(* IEC 61131-3 sources: Lasal-MCP/examples/SampleSource/LASALScreenAdvancedSolution/LASALScreenAdvancedSolution/LASALScreenAdvacnedSolution/Stations/Terminal/HMI/Class/DataRecordFileRead, 1 file *)

(* ---- DataRecordFileRead.st ---- *)
(*!
<Class
	Name               = "DataRecordFileRead"
	Revision           = "0.0"
	RealtimeTask       = "false"
	CyclicTask         = "false"
	BackgroundTask     = "true"
	DefBackground      = "10 ms"
	Sigmatek           = "false"
	OSInterface        = "false"
	HighPriority       = "false"
	Automatic          = "false"
	UpdateMode         = "Prescan"
	SharedCommandTable = "true"
	Objectsize         = "(444,120)">
	<Channels>
		<Server Name="IntError" Visualized="false" Initialize="false" WriteProtected="true" Retentive="false"/>
		<Server Name="ReadStep" Visualized="false" Initialize="false" WriteProtected="true" Retentive="false"/>
		<Server Name="StartRead" Visualized="true" Initialize="false" WriteProtected="false" Retentive="false"/>
		<Client Name="_FileSys" Required="false" Internal="false"/>
		<Client Name="_StdLib" Required="false" Internal="false"/>
		<Client Name="StringRAM" Required="true" Internal="false"/>
	</Channels>
</Class>
*)
DataRecordFileRead : CLASS
	TYPE
	  _READ_STEPS :  //! <Type Public="true" Name="_READ_STEPS"/>
	  (
	    RS_Idle,
	    RS_GetFileName,
	    RS_Open,
	    RS_WaitFileOpen,
	    RS_GetLength,
	    RS_WaitForGetLength,
	    RS_ReadFile,
	    RS_WaitForReadFile,
	    RS_CloseFile,
	    RS_WaitForClose,
	    RS_Error
	  )$UDINT;
	END_TYPE
  //Servers:
	ReadStep 	: SvrChCmd__READ_STEPS_PTofCls_DataRecordFileRead;
	IntError 	: SvrCh_DINT;
	StartRead 	: SvrCh_DINT;
  //Clients:
	_FileSys 	: CltChCmd__FileSys;
	_StdLib 	: CltChCmd__StdLib;
	StringRAM 	: CltChCmd_StringRAM;
  //Variables:
		FileName : ARRAY [0..99] OF CHAR;

		AsyncId 	: DINT;
		FileHandle 	: DINT;
		FileLength 	: UDINT;
		pReadData 	: ^DINT;
		FileIsRead 	: BOOL;
  //Functions:

	FUNCTION VIRTUAL GLOBAL Background
		VAR_INPUT
			EAX 	: UDINT;
		END_VAR
		VAR_OUTPUT
			state (EAX) 	: UDINT;
		END_VAR;

	FUNCTION GLOBAL ReadKoords
		VAR_INPUT
			pNoOfCoordinates 	: ^UDINT;
		END_VAR
		VAR_OUTPUT
			pCoord 	: ^_DOT;
		END_VAR;

	FUNCTION GLOBAL GetReadState
		VAR_OUTPUT
			IsRead 	: BOOL;
		END_VAR;

	FUNCTION GLOBAL SetReadState
		VAR_INPUT
			IsDrawing 	: BOOL;
		END_VAR;

	FUNCTION GLOBAL StartReading
		VAR_INPUT
			BufferSize 	: UDINT;
		END_VAR;
  //Tables:
	FUNCTION @STD
		VAR_OUTPUT
			ret_code	: CONFSTATES;
		END_VAR;
	FUNCTION GLOBAL TAB @CT_;
END_CLASS;

#pragma usingLtd _FileSys
#pragma usingLtd _StdLib
#pragma usingLtd StringRAM

FUNCTION VIRTUAL GLOBAL DataRecordFileRead::Background
	VAR_INPUT
		EAX 	: UDINT;
	END_VAR
	VAR_OUTPUT
		state (EAX) 	: UDINT;
	END_VAR
  VAR
  	stringLength : UDINT;
    asyncState : DINT;
    length : UDINT;
  END_VAR

  // ==========================================================================
  case ReadStep of

    // --------------------------------------------------------------
  	RS_Idle:

      if (StartRead = 1) then
         StartRead := 0;

         ReadStep := RS_GetFileName;
      end_if;

    // --------------------------------------------------------------
  	RS_GetFileName:

      stringLength := StringRAM.GetLength();

      StringRAM.GetDataAt(pData:= #FileName[0],
                          udSize:= stringLength,
                          udAt:= 0);

      ReadStep := RS_Open;

    // --------------------------------------------------------------
  	RS_Open:

      AsyncId := _FileSys.FileOpen_A(Async:= 1,
                                     filename:= #FileName[0],
                                     attributes:= ATT_READ_WRITE);

      ReadStep := RS_WaitFileOpen;

    // --------------------------------------------------------------
  	RS_WaitFileOpen:

      asyncState := _FileSys.GetAsyncState(ID:= to_udint(AsyncId),
                                           Erg:= #FileHandle);

      // ==================================================
      case asyncState of
        //---------------------------------------
        0:
          if (FileHandle >= 0) then
              ReadStep := RS_GetLength;
          else
            IntError := -1;
            ReadStep := RS_Error;
          end_if;

        //---------------------------------------
        RT_ERG_DELETED,
        RT_INVALID_ID:
          IntError := -2;
          ReadStep := RS_Error;

        //---------------------------------------
        RT_NOT_STARTED,
        RT_IN_PROGRESS:

      end_case;
      // ==================================================

    // --------------------------------------------------------------
  	RS_GetLength:

      AsyncId := _FileSys.FileLength_A(Async:= 1,
                                       handle:= FileHandle);
      ReadStep := RS_WaitForGetLength;

    // --------------------------------------------------------------
  	RS_WaitForGetLength:

      asyncState := _FileSys.GetAsyncState(ID:= to_udint(AsyncId),
                                           Erg:= #FileLength$dint);
        // ==================================================
      case asyncState of
        //---------------------------------------
        0:
          if (FileLength >= 0) then
            ReadStep := RS_ReadFile;
          end_if;

        //---------------------------------------
        RT_ERG_DELETED,
        RT_INVALID_ID:
            IntError := -3;
            ReadStep := RS_Error;

        //---------------------------------------
        RT_NOT_STARTED,
        RT_IN_PROGRESS:

      end_case;
     // ==================================================

    // --------------------------------------------------------------
  	RS_ReadFile:

      if (pReadData <> NIL) then
        _StdLib.Free(mptr:=pReadData);
      end_if;

      pReadData$^void := oc_StdLib.Malloc(size:= FileLength);

      AsyncId$UDINT := _FileSys.FileRead_A(Async:= 1,
                                           handle:= FileHandle,
                                           buffer:= pReadData,
                                           length:= FileLength);
      ReadStep := RS_WaitForReadFile;

    // --------------------------------------------------------------
  	RS_WaitForReadFile:

      asyncState := _FileSys.GetAsyncState(ID:= to_udint(AsyncId),
                                           Erg:= #FileHandle);
      // ==================================================
      case asyncState of
        //---------------------------------------
        0:
          if (length <> FileLength) then
            ReadStep := RS_CloseFile;
          else
            IntError := -4;
            ReadStep := RS_Error;
          end_if;

        //---------------------------------------
        RT_ERG_DELETED,
        RT_INVALID_ID:
          IntError := -5;
          ReadStep := RS_Error;

        //---------------------------------------
        RT_NOT_STARTED,
        RT_IN_PROGRESS:

        end_case;
       // ==================================================

    // --------------------------------------------------------------
  	RS_CloseFile:

      AsyncId := _FileSys.FileClose_A(Async:= 1,
                                      handle:= FileHandle);

      ReadStep := RS_WaitForClose;

    // --------------------------------------------------------------
  	RS_WaitForClose:

     asyncState := _FileSys.GetAsyncState(ID:= to_udint(AsyncId),
                                          Erg:= #FileHandle);

      // ==================================================
      case asyncState of
        //---------------------------------------
        0:
          if (FileHandle >= 0) then
            FileIsRead := TRUE;
            ReadStep := RS_Idle;
          else
            IntError := -6;
            ReadStep := RS_Error;
          end_if;
      end_case;
      // ==================================================

    // --------------------------------------------------------------
  	RS_Error:

  end_case;
  // ==========================================================================

	state := READY;

END_FUNCTION

FUNCTION GLOBAL DataRecordFileRead::ReadKoords
	VAR_INPUT
		pNoOfCoordinates 	: ^UDINT;
	END_VAR
	VAR_OUTPUT
		pCoord 	: ^_DOT;
	END_VAR

  pNoOfCoordinates^ := FileLength;
  pCoord := pReadData$^_DOT;

END_FUNCTION

FUNCTION GLOBAL DataRecordFileRead::GetReadState
	VAR_OUTPUT
		IsRead 	: BOOL;
	END_VAR

  IsRead := FileIsRead;

END_FUNCTION

FUNCTION GLOBAL DataRecordFileRead::SetReadState
	VAR_INPUT
		IsDrawing 	: BOOL;
	END_VAR

  FileIsRead := IsDrawing;

END_FUNCTION

FUNCTION GLOBAL DataRecordFileRead::StartReading
	VAR_INPUT
		BufferSize 	: UDINT;
	END_VAR

  if (pReadData <> NIL) then
    _StdLib.Free(mptr:=pReadData);
  end_if;

  pReadData$^void := _StdLib.Malloc(size:=BufferSize);

  if (pReadData <> NIL) then
      _StdLib.MemSet(dest:= pReadData,
                     value:= 0,
                     size:= BufferSize);
  end_if;

  ReadStep := RS_GetFileName;

END_FUNCTION
